PROGRAM MAIN
VAR
	sIPAddr			: STRING(15);
END_VAR

END_PROGRAM

(* stored: Version 1.1.0.1, ProductVersion 3.1.4024.9
   POU MAIN: Id {828f2a7a-e803-4f63-be04-ce2d692c8654}, SpecialFunc None *)
